Fanuc KAREL source: kt00706.KL

PROGRAM KT00706
%STACKSIZE=65535
%PRIORITY=65535
%NOLOCKGROUP
VAR
I1 : INTEGER
I2 : INTEGER
OUT : BOOLEAN
BEGIN
I1=2
I2=3
I1=2
I2=3
-- UNRESOLVED_PC line 12 opcodes [22 63 23] marker_code=64
END KT00706
